// TIA Portal V21 export
// export: Created 2026-10-23T21:22:24.3867133Z, ExportSetting WithReadOnly, DisplayName Totally Integrated Automation Portal, DisplayVersion V21 Update 1, DisplayName SINAMICS Startdrive Advanced, DisplayVersion V21 HF2, DisplayName SINAMICS Startdrive G110M, G120, G120C, G120D, G120P, G115D, DisplayVersion V21 HF2, DisplayName SINAMICS Startdrive G130, G150, S120, S150, G200, G220, S200, S210, S220, Innomotics MVD, DisplayVersion V21 HF2, DisplayName STEP 7 Professional, DisplayVersion V21 Update 1, DisplayName STEP 7 Safety, DisplayVersion V21, DisplayName Tech WebApplication, DisplayVersion V21, DisplayName WinCC Basic/Comfort/Advanced, DisplayVersion V21 Update 1, DisplayName WinCC Unified, DisplayVersion V21 Update 1
ORGANIZATION_BLOCK "OB_HwInterrupt"   // OB40, SCL, HardwareInterrupt
TITLE = Prozessalarm / Hardware interrupt
{ S7_Optimized_Access := 'TRUE' }
// Minimaler Prozessalarm-OB / Minimal hardware interrupt OB
// stored: AutoNumber false, CodeModifiedDate 2026-10-23T19:38:38.9967876Z, CompileDate 2026-10-23T19:38:38.9967876Z, ConstantName OB_OB_HwInterrupt, CreationDate 2026-10-23T19:38:17.2685443Z, DownloadDate 0001-01-01T00:00:00Z, EventClass Hardware interrupt, InterfaceModifiedDate 2008-07-21T16:55:29.2443395Z, IsConsistent true, LoadMemoryLength 3693, ModifiedDate 2026-10-23T19:38:38.9967876Z, ParameterModified 2008-07-21T16:55:29.2443395Z, ProcessImagePartNumber 65535, SetENOAutomatically false, StructureModified 2008-07-21T16:55:29.2443395Z, WorkMemoryLength 120
   VAR_INPUT
      LADDR : HW_IO;   // Hardware identifier
      USI : Word;   // User structure identifier
      IChannel : USInt;   // Interrupt channel number
      EventType : Byte;   // EventType
      PointAddr : DWord;
   END_VAR
BEGIN

       // Count hardware interrupts
       "DB_Machine".TotalCountUnsigned := "DB_Machine".TotalCountUnsigned + 1;
END_ORGANIZATION_BLOCK
